// TIA Portal V20 export
// export: Created 2026-10-20T12:45:14.8946516Z, ExportSetting WithDefaults, DisplayName Totally Integrated Automation Portal, DisplayVersion V20 Update 6, DisplayName TIA Portal Openness, DisplayVersion V20 Update 6, DisplayName TIA Portal Version Control Interface, DisplayVersion V20 Update 6, DisplayName SINAMICS Startdrive Advanced, DisplayVersion V20 SP1, DisplayName SINAMICS Startdrive G130, G150, S120, S150, SINAMICS MV, G220, S200, S210, DisplayVersion V20 SP1, DisplayName SINAMICS Startdrive G110M, G120, G120C, G120D, G120P, G115D, DisplayVersion V20 SP1, DisplayName STEP 7 Professional, DisplayVersion V20 Update 6, DisplayName STEP 7 Safety, DisplayVersion V20 Update 2, DisplayName WinCC Basic/Comfort/Advanced, DisplayVersion V20 Update 6, DisplayName WinCC Unified, DisplayVersion V20 Update 6
FUNCTION "Feed_ECNV" : Void   // FC1, SCL
{ S7_Optimized_Access := 'TRUE' }
VERSION : 0.1
// stored: AutoNumber true, IsIECCheckEnabled false, SetENOAutomatically false, UDAEnableTagReadback false
   VAR_INPUT
      System_No : UInt;
      Safety_OK : Bool;
      Overhang_Left : Bool;
      Overhang_Right : Bool;
   END_VAR
   VAR_IN_OUT
      System_Busy : Bool;
   END_VAR
BEGIN
   //Sensors
   "HMI_CNV_Left" := "Control_DB".ECnv_Sys[#System_No].Inputs.Left;
   "HMI_CNV_Lpd1" := "Control_DB".ECnv_Sys[#System_No].Inputs.Lpd1;
   "HMI_CNV_Lpd2" := "Control_DB".ECnv_Sys[#System_No].Inputs.Center;
   "HMI_CNV_Rpd1" := "Control_DB".ECnv_Sys[#System_No].Inputs.Rpd1;
   "HMI_CNV_Right" := "Control_DB".ECnv_Sys[#System_No].Inputs.Right;

   "HMI_CNV_Sdetect1" := #Overhang_Left;
   "HMI_CNV_Sdetect2" := #Overhang_Right;

   //Feedback
   "Mode_HMI" := "Control_DB".ECnv_Sys[#System_No].Mode;
   "Enabled_HMI" := "Control_DB".ECnv_Sys[#System_No].Enabled;
   "Error_HMI" := "Control_DB".ECnv_Sys[#System_No].Error;
   "Warning_HMI" := "Control_DB".ECnv_Sys[#System_No].Warning;
   "Stopped_HMI" := "Control_DB".ECnv_Sys[#System_No].Stopped;
   "Running_HMI" := "Control_DB".ECnv_Sys[#System_No].Running;
   "Ready_For_Task_HMI" := "Control_DB".ECnv_Sys[#System_No].Ready_For_Task;
   "Cnv_Occupied_HMI" := "Control_DB".ECnv_Sys[#System_No].Cnv_Occupied;
   "Shuttle_in_place_HMI" := "Control_DB".ECnv_Sys[#System_No].Shuttle_In_Place;
   "Current_Task_Type_HMI" := "Control_DB".ECnv_Sys[#System_No].Current_Task_Type;
   "Current_Task_ID_HMI" := "Control_DB".ECnv_Sys[#System_No].Current_Task_ID;
   "SM_State_HMI" := "Control_DB".ECnv_Sys[#System_No].SM_State;
   "Pallet_Type_HMI" := "Control_DB".ECnv_Sys[#System_No].Pallet_Type;
   IF "Control_DB".ECnv_Sys[#System_No].Motor.Forward THEN
       "Motor_Direction_HMI" := 1;
   ELSIF "Control_DB".ECnv_Sys[#System_No].Motor.Reverse THEN
       "Motor_Direction_HMI" := 2;
   ELSE
       "Motor_Direction_HMI" := 0;
   END_IF;
   "Motor_Speed_Requested_HMI" := "Control_DB".ECnv_Sys[#System_No].Motor.Speed;
   "Motor_Speed_Actual_HMI" := "Control_DB".ECnv_Sys[#System_No].Motor.Speed_Actual;
   "CNV_Motor_Ready" := "Control_DB".ECnv_Sys[#System_No].Motor.Ready;
   "CNV_Motor_Current_Actual_HMI" := "Control_DB".ECnv_Sys[#System_No].Motor.Actual_Current;
   "CNV_Motor_Actual_Torque" := "Control_DB".ECnv_Sys[#System_No].Motor.Actual_Torque;
   "Transfer_To_ID_HMI" := "Control_DB".ECnv_Sys[#System_No].Instruction.Transfer_To_ID;
   "Transfer_From_ID_HMI" := "Control_DB".ECnv_Sys[#System_No].Instruction.Transfer_From_ID;

   IF "Control_DB".ECnv_Sys[#System_No].Motor.Error THEN
       "CNV_Motor_Status_HMI" := 2;
   ELSIF "Control_DB".ECnv_Sys[#System_No].Motor.Enabled THEN
       "CNV_Motor_Status_HMI" := 1;
   ELSIF NOT "Control_DB".ECnv_Sys[#System_No].Motor.Enabled THEN
       "CNV_Motor_Status_HMI" := 0;
   END_IF;

   "Safety_OK_HMI" := #Safety_OK;

   //Instructions
   IF ("HMI_Box_Connected_1" = #System_No OR ("HMI_Box_Connected_1" >= (#System_No * 10) + 1 AND "HMI_Box_Connected_1" <= (#System_No * 10) + 8)) OR
       ("HMI_Box_Connected_2" = #System_No OR ("HMI_Box_Connected_1" >= (#System_No * 10) + 1 AND "HMI_Box_Connected_1" <= (#System_No * 10) + 8))
   THEN
       #System_Busy := TRUE;
   ELSE
       #System_Busy := FALSE;
       "Control_DB".ECnv_Sys[#System_No].Instruction.Stop := "Stop_HMI";
       "Control_DB".ECnv_Sys[#System_No].Instruction.Execute := "Manual_Fwd_HMI" OR "Manual_Bwd_HMI";
       IF "BT_Confirmation_HMI" THEN
           "Control_DB".VTD_Sys[#System_No].Instruction.Mode_Change :=
           "Control_DB".ECnv_Sys[#System_No].Instruction.Mode_Change :=
           "Control_DB".LCnv_Sys[#System_No].Cnv_Level[1].Cnv1.Instruction.Mode_Change :=
           "Control_DB".LCnv_Sys[#System_No].Cnv_Level[2].Cnv1.Instruction.Mode_Change :=
           "Control_DB".LCnv_Sys[#System_No].Cnv_Level[3].Cnv1.Instruction.Mode_Change :=
           "Control_DB".LCnv_Sys[#System_No].Cnv_Level[4].Cnv1.Instruction.Mode_Change :=
           "Control_DB".LCnv_Sys[#System_No].Cnv_Level[5].Cnv1.Instruction.Mode_Change :=
           "Control_DB".LCnv_Sys[#System_No].Cnv_Level[6].Cnv1.Instruction.Mode_Change :=
           "Control_DB".LCnv_Sys[#System_No].Cnv_Level[7].Cnv1.Instruction.Mode_Change :=
           "Control_DB".LCnv_Sys[#System_No].Cnv_Level[8].Cnv1.Instruction.Mode_Change :=
           "Control_DB".LCnv_Sys[#System_No].Cnv_Level[1].Cnv2.Instruction.Mode_Change :=
           "Control_DB".LCnv_Sys[#System_No].Cnv_Level[2].Cnv2.Instruction.Mode_Change :=
           "Control_DB".LCnv_Sys[#System_No].Cnv_Level[3].Cnv2.Instruction.Mode_Change :=
           "Control_DB".LCnv_Sys[#System_No].Cnv_Level[4].Cnv2.Instruction.Mode_Change :=
           "Control_DB".LCnv_Sys[#System_No].Cnv_Level[5].Cnv2.Instruction.Mode_Change :=
           "Control_DB".LCnv_Sys[#System_No].Cnv_Level[6].Cnv2.Instruction.Mode_Change :=
           "Control_DB".LCnv_Sys[#System_No].Cnv_Level[7].Cnv2.Instruction.Mode_Change :=
           "Control_DB".LCnv_Sys[#System_No].Cnv_Level[8].Cnv2.Instruction.Mode_Change := "Mode_Change_HMI";
           "Mode_Change_HMI(1)" := "Mode_Change_HMI";
           "BT_Confirmation_HMI" := FALSE;
       END_IF;

       "Control_DB".ECnv_Sys[#System_No].Instruction.Enable := "Enable_HMI";

       "Control_DB".ECnv_Sys[#System_No].Instruction.Reset := "Reset_HMI" OR "Reset_All" OR
       "Screen_DB_1".Reset_All[1] OR "CNV_HMI".Reset[1] OR
       "Screen_DB_1".Reset_All[2] OR "CNV_HMI".Reset[2];

       IF "Control_DB".ECnv_Sys[#System_No].Mode <> 3 THEN
           "Control_DB".ECnv_Sys[#System_No].Instruction.Foward := "Manual_Fwd_HMI";
           "Control_DB".ECnv_Sys[#System_No].Instruction.Backward := "Manual_Bwd_HMI";
           "Control_DB".ECnv_Sys[#System_No].Instruction.Start_Transfer := "Start_Transfer_HMI";
           IF "Control_DB".ECnv_Sys[#System_No].Mode = 1 THEN
               "Control_DB".ECnv_Sys[#System_No].Instruction.Start_Transfer_Backward := "Transfer_Backward";
           END_IF;
           "Control_DB".ECnv_Sys[#System_No].Instruction.Task_ID := "Task_ID_HMI";
           "Control_DB".ECnv_Sys[#System_No].Instruction.Pallet_Align_Left := "Pallet_Align_Left_HMI";
           "Control_DB".ECnv_Sys[#System_No].Instruction.Pallet_Align_Right := "Pallet_Align_Right_HMI";
           "Control_DB".ECnv_Sys[#System_No].Instruction.Pallet_Align_Center := "Pallet_Align_Center_HMI";
           IF "Mode_Change_HMI" <> 2 THEN
               "Control_DB".ECnv_Sys[#System_No].Instruction.Pallet_Allignment := "Pallet_Allignment_HMI" := FALSE;
           ELSE
               "Control_DB".ECnv_Sys[#System_No].Instruction.Pallet_Allignment := "Pallet_Allignment_HMI";
           END_IF;
           IF "CNV_HMI".In_Out[#System_No] THEN // 0 = ECNV RECEIVE, 1 = ECONV SEND
               "Control_DB".ECnv_Sys[#System_No].Instruction.Transfer_To_ID := "CNV_ID_HMI(1)";
               "Control_DB".ECnv_Sys[#System_No].Instruction.Transfer_From_ID := 0;
           ELSE
               "Control_DB".ECnv_Sys[#System_No].Instruction.Transfer_To_ID := 0;
               "Control_DB".ECnv_Sys[#System_No].Instruction.Transfer_From_ID := "CNV_ID_HMI(1)";
           END_IF;
       END_IF;
   END_IF;
END_FUNCTION
